Fanuc KAREL source: kx00030.KL

PROGRAM KX00030
%STACKSIZE=65535
%PRIORITY=65535
VAR
I : INTEGER
J : INTEGER
B : BOOLEAN
F : FILE
S : STRING[80]
P : XYZWPR
BEGIN
I=1
END KX00030
